(* IEC 61131-3 sources: PLC-Static-Analysis/modules/plc-rules/src/test/resources/PLCA-P003/global, 1 file *)

(* ---- two.st ---- *)
VAR_GLOBAL
    gfbPulse : TP;
END_VAR

PROGRAM P_A
gfbPulse(IN := TRUE, PT := T#1S);
END_PROGRAM

PROGRAM P_B
gfbPulse(IN := TRUE, PT := T#2S); // PLCA-P003
END_PROGRAM
